// TIA Portal V21 export
Screen "R10_LampA"  1024x768, Number=50, Template=Tpl
  ScreenLayer 
    Rectangle "P_LampAlarm" at 10,10 size 100x30
      RangeAppearanceAnimation "RangeAppearanceAnimation"
        tag P_SwOn
        0..0: back #aaaaaa, fore #000000
        1..1: back #dc0000, fore #000000, flashing
